(* IEC 61131-3 sources: plcassist-cli/packages/volt-lsp-iec/test-corpus/awa-palletizer/Device/Plc Logic/Application/Library Manager/L_UM1P_MulticoreBasic, 31 files *)

(* ---- L_UM1P_CONSTANTS.gvl ---- *)
VAR_GLOBAL
	C_UNDEFTASKINDEX : INT := -1;
	C_BITMASKTASKID : UDINT := UDINT#16#FF;
	C_MAXCORES : UINT := 4;
	C_MAXSYNCTASKS : UINT := 3;
END_VAR

(* ---- L_UM1P_INTERNAL.gvl ---- *)
VAR_GLOBAL
	BASICINFRASTRUCTURE : L_UM1P_BasicInfrastructure;
	C_MAXTASK : WORD := 31;
	C_MAXADDSYNCTASKS : WORD := 3;
	CDIENUMSTARTVALUE : DINT := 90000;
END_VAR

(* ---- L_UM1P_IBARRIER.itf ---- *)
INTERFACE L_UM1P_IBARRIER
END_INTERFACE

METHOD QUERYBARRIER
VAR_INPUT
	DWBARRIERID : DWORD;
END_VAR
END_METHOD

(* ---- L_UM1P_IFUNCTIONCALL.itf ---- *)
INTERFACE L_UM1P_IFUNCTIONCALL
END_INTERFACE

METHOD CALL
VAR_INPUT
	PINPUTDATA : POINTER TO BYTE;
	POUTPUTDATA : POINTER TO BYTE;
END_VAR
END_METHOD

(* ---- L_UM1P_IMCCALL.itf ---- *)
INTERFACE L_UM1P_IMCCALL
END_INTERFACE

METHOD CALLFUNCTION
VAR_INPUT
	UIINPUTDATAIDX : UINT;
	UIOUTPUTDATAIDX : UINT;
END_VAR
END_METHOD

METHOD COPYINPUTS : BOOL
VAR_INPUT
	IDX : WORD;
END_VAR
END_METHOD

METHOD COPYOUTPUTS : BOOL
VAR_INPUT
	IDX : WORD;
END_VAR
END_METHOD

METHOD FUNCTIONWASCALLEDTWICE : BOOL
VAR_INPUT
	IDX : WORD;
END_VAR
END_METHOD

METHOD HANDLESTANDARDCALL : BOOL
END_METHOD

METHOD SYNCOUTPUTS
VAR_INPUT
	UICOPYOUTPUTFROMIDX : UINT;
	UICOPYOUTPUTTOIDX : UINT;
END_VAR
END_METHOD

(* ---- L_UM1P_IMCCALLINFO.itf ---- *)
INTERFACE L_UM1P_IMCCALLINFO
END_INTERFACE

(* ---- L_UM1P_ISETPOINTINFO.itf ---- *)
INTERFACE L_UM1P_ISETPOINTINFO
END_INTERFACE

(* ---- L_UM1P_ISYNCPOINTCLIENT.itf ---- *)
INTERFACE L_UM1P_ISYNCPOINTCLIENT
END_INTERFACE

(* ---- L_UM1P_ISYNCPOINTSERVER.itf ---- *)
INTERFACE L_UM1P_ISYNCPOINTSERVER
END_INTERFACE

METHOD SUBSCRIBE : DWORD
VAR_INPUT
	ITFCLIENT : L_UM1P_ISyncPointClient;
END_VAR
END_METHOD

(* ---- L_UM1P_MULTICOREDATASENDER.itf ---- *)
INTERFACE L_UM1P_MULTICOREDATASENDER
END_INTERFACE

METHOD UPDATEINPUTDATA : BOOL
VAR_INPUT
	PTRAGET : POINTER TO BYTE;
	DISIZE : DINT;
	ETYPE : TYPE_CLASS;
END_VAR
END_METHOD

(* ---- GETBOOLEANPROPERTY.fun ---- *)
FUNCTION GETBOOLEANPROPERTY : BOOL
VAR_INPUT
	STKEY : WSTRING;
END_VAR
END_FUNCTION

(* ---- GETCOMPANY.fun ---- *)
FUNCTION GETCOMPANY : WSTRING
END_FUNCTION

(* ---- GETNUMBERPROPERTY.fun ---- *)
FUNCTION GETNUMBERPROPERTY : DINT
VAR_INPUT
	STKEY : WSTRING;
END_VAR
END_FUNCTION

(* ---- GETTEXTPROPERTY.fun ---- *)
FUNCTION GETTEXTPROPERTY : WSTRING
VAR_INPUT
	STKEY : WSTRING;
END_VAR
END_FUNCTION

(* ---- GETTEXTPROPERTY2.fun ---- *)
FUNCTION GETTEXTPROPERTY2 : POINTER TO WSTRING
VAR_INPUT
	STKEY : WSTRING;
END_VAR
END_FUNCTION

(* ---- GETTITLE.fun ---- *)
FUNCTION GETTITLE : WSTRING
END_FUNCTION

(* ---- GETVERSION.fun ---- *)
FUNCTION GETVERSION : VERSION
END_FUNCTION

(* ---- GETVERSIONPROPERTY.fun ---- *)
FUNCTION GETVERSIONPROPERTY : VERSION
VAR_INPUT
	STKEY : WSTRING;
END_VAR
END_FUNCTION

(* ---- L_SSYP_TASKISSYNCHRONIZED.fun ---- *)
FUNCTION L_SSYP_TASKISSYNCHRONIZED : BOOL
VAR_INPUT
	PTASKDESC : POINTER TO Task_Desc2;
END_VAR
END_FUNCTION

(* ---- L_UM1P_GETCURRENTTASKINDEX.fun ---- *)
FUNCTION L_UM1P_GETCURRENTTASKINDEX : INT
END_FUNCTION

(* ---- L_UM1P_INSERTFUNCTIONCALL.fun ---- *)
FUNCTION L_UM1P_INSERTFUNCTIONCALL : L_IE1P_Error
VAR_INPUT
	TASKID : INT;
	FUNCTIONCALLTOADD : POINTER TO L_UM1P_CallStackInfo;
END_VAR
END_FUNCTION

(* ---- L_UM1P_ISCALLEDINIDENTICALTASK.fun ---- *)
FUNCTION L_UM1P_ISCALLEDINIDENTICALTASK : BOOL
VAR_INPUT
	ICALLCYCLEREFERENCE : INT;
END_VAR
END_FUNCTION

(* ---- L_UM1P_ISCALLEDINMOTIONTASK.fun ---- *)
FUNCTION L_UM1P_ISCALLEDINMOTIONTASK : BOOL
VAR_INPUT
	TASKINDEX : INT;
END_VAR
VAR_OUTPUT
	DWCALLCYCLE : DWORD;
END_VAR
END_FUNCTION

(* ---- GLOBALTEXTLIST.fb ---- *)
FUNCTION_BLOCK GLOBALTEXTLIST
VAR
	M_TEXTLISTFILE : STRING(255);
	_STNAMESPACE : STRING;
END_VAR
END_FUNCTION_BLOCK

(* ---- L_UM1P_BASICINFRASTRUCTURE.fb ---- *)
FUNCTION_BLOCK L_UM1P_BASICINFRASTRUCTURE
VAR_INPUT
	ACALLSTACK : ARRAY [0..L_UM1P_Internal.c_MaxTask] OF L_UM1P_CallStack;
END_VAR
VAR_OUTPUT
	TASKSYNCAVAILABLE : ARRAY [0..L_UM1P_Internal.c_MaxTask] OF INT := [L_UM1P_Internal.c_MaxTask(-1)];
	TASKCYCLETIME : ARRAY [0..L_UM1P_Internal.c_MaxTask] OF DWORD;
END_VAR
VAR
	_HEVENTRESETDONE : RTS_IEC_HANDLE := RTS_INVALID_HANDLE;
	_HINTERFACERESETDONE : RTS_IEC_HANDLE := RTS_INVALID_HANDLE;
	_HEVENTDOWNLOADDONE : RTS_IEC_HANDLE := RTS_INVALID_HANDLE;
	_HINTERFACEDOWNLOADDONE : RTS_IEC_HANDLE := RTS_INVALID_HANDLE;
	_HEVENTBRI : RTS_IEC_HANDLE := SysTypes.RTS_INVALID_HANDLE;
	_HINTERFACEBRI : RTS_IEC_HANDLE := SysTypes.RTS_INVALID_HANDLE;
	_HEVENTBWO_ENTRY : RTS_IEC_HANDLE := SysTypes.RTS_INVALID_HANDLE;
	_HINTERFACEBWO_ENTRY : RTS_IEC_HANDLE := SysTypes.RTS_INVALID_HANDLE;
	BUSCYCLETASKID : UDINT := 16#FFFFFFFF;
	SYNCTASKID : ARRAY [1..L_UM1P_Internal.c_MaxAddSyncTasks] OF UDINT := [L_UM1P_Internal.c_MaxAddSyncTasks(16#FFFFFFFF)];
	ISYNCTASKCOUNT : INT := 0;
	DWCALL1 : DWORD;
	DWCALL2 : DWORD;
	APPCOUNT : DWORD;
	TASKCOUNT : DWORD;
	SINSTANCESTRFULL : STRING(255);
	SZAPPLICATION : STRING := '';
END_VAR
END_FUNCTION_BLOCK

METHOD EVENTCALLBACK : RTS_IEC_RESULT
VAR_INPUT
	PEVENTPARAM : POINTER TO EventParam;
END_VAR
END_METHOD

METHOD GETAPPNAME : STRING
END_METHOD

METHOD METH : BOOL
END_METHOD

METHOD REGISTEREVENTS
VAR_INPUT
	XONLYCALLBACKFUNCTION : BOOL;
END_VAR
END_METHOD

METHOD REGISTERMOTIONFUNCTION : BOOL
VAR_INPUT
	TASKINDEX : INT;
END_VAR
END_METHOD

METHOD UNREGISTEREVENTS
VAR_INPUT
	XONLYCALLBACKFUNCTION : BOOL;
END_VAR
END_METHOD

METHOD FB_EXIT : BOOL
VAR_INPUT
	BINCOPYCODE : BOOL;
END_VAR
END_METHOD

METHOD FB_INIT : BOOL
VAR_INPUT
	BINITRETAINS : BOOL;
	BINCOPYCODE : BOOL;
END_VAR
END_METHOD

METHOD FB_REINIT : BOOL
END_METHOD

(* ---- L_UM1P_CALLSTACK.fb ---- *)
FUNCTION_BLOCK L_UM1P_CALLSTACK
VAR_OUTPUT
	XNOTCALLED : BOOL;
END_VAR
VAR
	PRES1 : RTS_IEC_RESULT;
	HSEMFILLSTACK : RTS_IEC_HANDLE;
	WVALIDSTACK : WORD;
	ALASTENTRY : ARRAY [1..2] OF POINTER TO L_UM1P_CallStackInfo;
	AFIRSTENTRY : ARRAY [1..2] OF POINTER TO L_UM1P_CallStackInfo;
	PACTENTRY : POINTER TO L_UM1P_CallStackInfo;
	IDX : WORD;
	DWSETCYCLECOUNTER : DWORD;
	DWACTCYCLECOUNTER : DWORD;
END_VAR
END_FUNCTION_BLOCK

METHOD INSERTFUNCTIONCALL : BOOL
VAR_INPUT
	FUNCTIONCALLTOADD : POINTER TO L_UM1P_CallStackInfo;
END_VAR
END_METHOD

METHOD SWITCH : BOOL
END_METHOD

METHOD FB_EXIT : BOOL
VAR_INPUT
	BINCOPYCODE : BOOL;
END_VAR
END_METHOD

METHOD FB_INIT : BOOL
VAR_INPUT
	BINITRETAINS : BOOL;
	BINCOPYCODE : BOOL;
END_VAR
END_METHOD

METHOD FB_REINIT : BOOL
END_METHOD

(* ---- L_UM1P_DATARECEIVER.fb ---- *)
FUNCTION_BLOCK L_UM1P_DATARECEIVER
VAR_INPUT
	ITFDATASENDER : L_UM1P_MultiCoreDataSender;
	ANYMIRROR : __SYSTEM.AnyType;
END_VAR
VAR_OUTPUT
	XVALID : BOOL;
END_VAR
VAR
	_HMYIECTASK : RTS_IEC_HANDLE;
	_XINITDONE : BOOL;
	_FBCYCLICCALLER : L_UBUP_CyclicCaller;
	_XCALLBRI : BOOL;
END_VAR
END_FUNCTION_BLOCK

METHOD AFTERWRITEOUTPUTS : INT
END_METHOD

METHOD BEFOREREADINPUTS : INT
END_METHOD

METHOD UPDATEMIRRORDATA : BOOL
END_METHOD

(* ---- L_UM1P_DATASENDER.fb ---- *)
FUNCTION_BLOCK L_UM1P_DATASENDER
VAR_INPUT
	ANYSOURCE : __SYSTEM.AnyType;
END_VAR
VAR
	_HMYIECTASK : RTS_IEC_HANDLE;
	_XINITDONE : BOOL;
	ISBUSTASK : BOOL;
	UIOSHANDLE : RTS_IEC_HANDLE;
END_VAR
END_FUNCTION_BLOCK

METHOD REQUESTINTERFACE : BOOL
VAR_INPUT
	ID : DINT;
	PITFUNKNOWN : POINTER TO L_UBUP.L_UBUP_IUnknown;
END_VAR
END_METHOD

METHOD UPDATEINPUTDATA : BOOL
VAR_INPUT
	PTRAGET : POINTER TO BYTE;
	DISIZE : DINT;
	ETYPE : TYPE_CLASS;
END_VAR
END_METHOD

(* ---- L_UM1P_MCCALL.fb ---- *)
FUNCTION_BLOCK L_UM1P_MCCALL
VAR_INPUT
	ICALLCYCLEREFERENCE : INT;
	ITFMCCALL : L_UM1P_IMCCall;
END_VAR
VAR_OUTPUT
	XERROR : BOOL;
	EERRORID : L_IE1P_Error;
	XMCHANDLINGACTIVE : BOOL;
	C_BUFFERDEPTHINPUT : WORD := 2;
	C_BUFFERDEPTHOUTPUT : WORD := 2;
END_VAR
VAR
	CALLSTACKINFO1 : ARRAY [1..c_BufferDepthInput] OF L_UM1P_CallStackInfo;
	DWCALLCYCLE : DWORD;
	DWCALLCYCLETMP : DWORD;
	XMIRROR : BOOL;
	IDX : WORD;
	LASTIDX : WORD := 1;
END_VAR
END_FUNCTION_BLOCK

METHOD ISCALLEDINIDENTICALTASK : BOOL
VAR_INPUT
	ICALLCYCLEREFERENCE : INT;
END_VAR
END_METHOD

(* ---- L_UM1P_MCMULTIPLECALL.fb ---- *)
FUNCTION_BLOCK L_UM1P_MCMULTIPLECALL
VAR_INPUT
	ICALLCYCLEREFERENCE : INT;
	ITFMCCALL : L_UM1P_IMCCall;
END_VAR
VAR_OUTPUT
	XERROR : BOOL;
	EERRORID : L_IE1P_Error;
	C_BUFFERDEPTHINPUT : WORD := 4;
	C_BUFFERDEPTHOUTPUT : WORD := 2;
END_VAR
VAR
	CALLSTACKINFO1 : ARRAY [1..c_BufferDepthInput] OF L_UM1P_CallStackInfo;
	DWCALLCYCLE : DWORD;
	DWCALLCYCLE2ND : DWORD;
	DWCALLCYCLETMP : DWORD;
	XMIRROR : BOOL;
	IDX : WORD;
	IDX2NDCALL : WORD;
	LASTIDX : WORD := 1;
END_VAR
END_FUNCTION_BLOCK

METHOD ISCALLEDINIDENTICALTASK : BOOL
VAR_INPUT
	ICALLCYCLEREFERENCE : INT;
END_VAR
END_METHOD

(* ---- L_UM1P_MEMMAPPING.fb ---- *)
FUNCTION_BLOCK L_UM1P_MEMMAPPING
VAR_INPUT
	PSRC : POINTER TO BYTE;
	PDEST : POINTER TO BYTE;
	DWSIZE : DWORD;
END_VAR
VAR
	_CYCLICCALLER : L_UBUP_CyclicCaller;
END_VAR
END_FUNCTION_BLOCK

METHOD BEFOREREADINPUTS : INT
END_METHOD
